SUBAPPLICATION doppeltwirkend (* Subapplication Type *)
  (* Standard: 61499-2 *)
  (* Version 1.0, 2023-01-29, Franz *)
  IMPORT DataPanel::io::MI::DQ::DataPanel_MI_DO::Invalid;
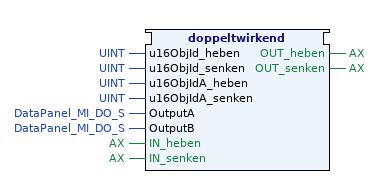
  VAR_INPUT
    u16ObjId_heben : UINT;
    u16ObjId_senken : UINT;
    u16ObjIdA_heben : UINT;
    u16ObjIdA_senken : UINT;
    OutputA : DataPanel::io::MI::DQ::DataPanel_MI_DO_S := Invalid;
    OutputB : DataPanel::io::MI::DQ::DataPanel_MI_DO_S := Invalid;
  END_VAR
  SOCKETS
    IN_heben : adapter::types::unidirectional::AX;
    IN_senken : adapter::types::unidirectional::AX;
  END_SOCKETS
  PLUGS
    OUT_heben : adapter::types::unidirectional::AX;
    OUT_senken : adapter::types::unidirectional::AX;
  END_PLUGS
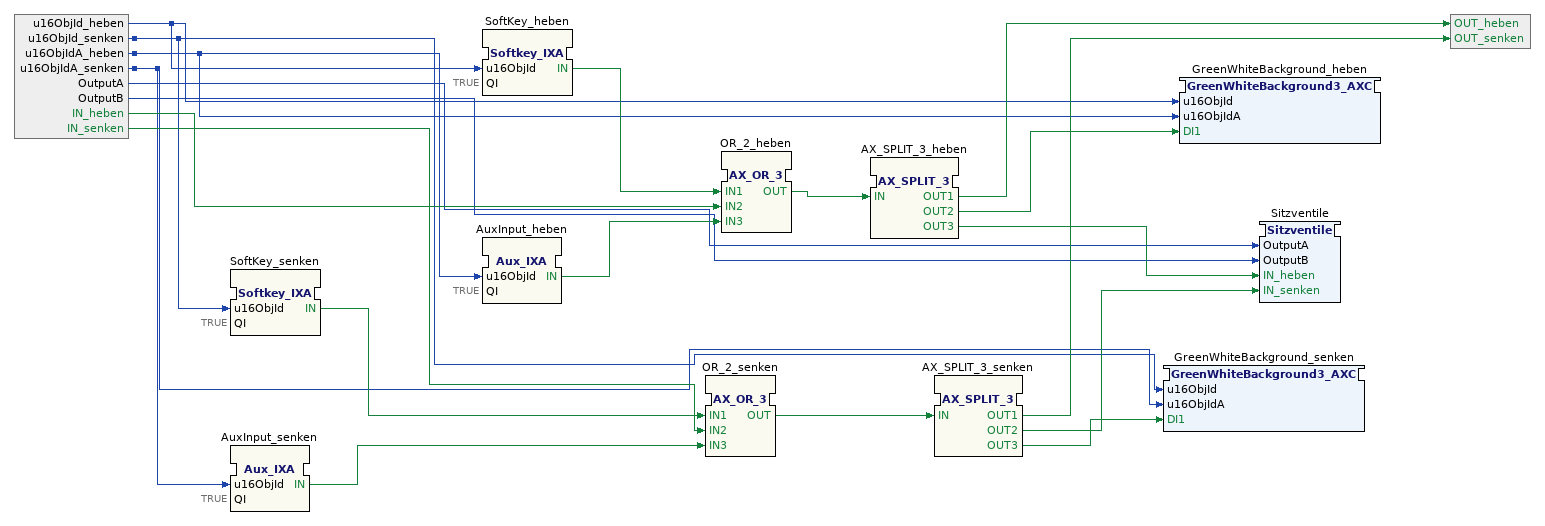
  FBS
    OR_2_heben : adapter::booleanOperators::AX_OR_3;
    AX_SPLIT_3_heben : adapter::events::unidirectional::AX_SPLIT_3;
    OR_2_senken : adapter::booleanOperators::AX_OR_3;
    AX_SPLIT_3_senken : adapter::events::unidirectional::AX_SPLIT_3;
    SoftKey_heben : isobus::UT::io::Softkey::Softkey_IXA(QI := TRUE);
    AuxInput_heben : isobus::UT::io::Auxiliary::IN::Aux_IXA(QI := TRUE);
    SoftKey_senken : isobus::UT::io::Softkey::Softkey_IXA(QI := TRUE);
    AuxInput_senken : isobus::UT::io::Auxiliary::IN::Aux_IXA(QI := TRUE);
  END_FBS
  SUBAPPS
    GreenWhiteBackground_heben : MyLib::sys::GreenWhiteBackground3_AXC;
    GreenWhiteBackground_senken : MyLib::sys::GreenWhiteBackground3_AXC;
    Sitzventile : Sitzventile;
  END_SUBAPPS
  DATA_CONNECTIONS
    OutputB TO Sitzventile.OutputB;
    OutputA TO Sitzventile.OutputA;
    u16ObjIdA_senken TO AuxInput_senken.u16ObjId;
    u16ObjIdA_heben TO AuxInput_heben.u16ObjId;
    u16ObjId_heben TO SoftKey_heben.u16ObjId;
    u16ObjId_senken TO SoftKey_senken.u16ObjId;
    u16ObjId_heben TO GreenWhiteBackground_heben.u16ObjId;
    u16ObjId_senken TO GreenWhiteBackground_senken.u16ObjId;
    u16ObjIdA_heben TO GreenWhiteBackground_heben.u16ObjIdA;
    u16ObjIdA_senken TO GreenWhiteBackground_senken.u16ObjIdA;
  END_CONNECTIONS
  ADAPTER_CONNECTIONS
    SoftKey_heben.IN TO OR_2_heben.IN1;
    IN_heben TO OR_2_heben.IN2;
    AuxInput_heben.IN TO OR_2_heben.IN3;
    OR_2_heben.OUT TO AX_SPLIT_3_heben.IN;
    AX_SPLIT_3_heben.OUT1 TO OUT_heben;
    AX_SPLIT_3_heben.OUT2 TO GreenWhiteBackground_heben.DI1;
    AX_SPLIT_3_heben.OUT3 TO Sitzventile.IN_heben;
    SoftKey_senken.IN TO OR_2_senken.IN1;
    IN_senken TO OR_2_senken.IN2;
    AuxInput_senken.IN TO OR_2_senken.IN3;
    OR_2_senken.OUT TO AX_SPLIT_3_senken.IN;
    AX_SPLIT_3_senken.OUT1 TO OUT_senken;
    AX_SPLIT_3_senken.OUT2 TO Sitzventile.IN_senken;
    AX_SPLIT_3_senken.OUT3 TO GreenWhiteBackground_senken.DI1;
  END_CONNECTIONS
END_SUBAPPLICATION
